(* IEC 61131-3 sources: Caravan/Archiv/12-04-19/Stations/Terminal/HMI/Network, 1 file *)

(* ---- ConfigObjects.st ---- *)
FUNCTION GLOBAL TAB TASK_CONF
_K_TASK, _K_REAL,
_K_END_VAR,

_K_TASK, _K_CYCLIC,
_K_END_VAR,

_K_TASK, _K_BACKGROUND,
_K_END_VAR,

_K_END_CONF
END_FUNCTION

FUNCTION GLOBAL TAB IPR_CONF
_K_IPR
	0$UINT,
_K_END_VAR,
_K_END_CONF
END_FUNCTION

FUNCTION GLOBAL TAB CONFIG_TABLES
00081$UINT,
0$UINT, 0, 10, "_ALARMDISPLAY",
0$UINT, 0, 11, "_ALARMX0PARA",
0$UINT, 0, 2, "_ALARMX1PARA",
0$UINT, 0, 19, "_ALARMXBUFFER",
0$UINT, 0, 1, "_BIT32",
0$UINT, 0, 1, "_BIT32RAM",
0$UINT, 0, 4, "_CAN",
0$UINT, 1, 3, "_CHECKONLINESTATUS",
0$UINT, 1, 0, "_CHECKSUM",
0$UINT, 1, 19, "_FILESYS",
0$UINT, 0, 14, "_GLOBAL",
0$UINT, 1, 2, "_GRAFIX",
0$UINT, 0, 1, "_HOTALARM",
0$UINT, 1, 8, "_IP",
0$UINT, 1, 1, "_IPCONFIGIF",
0$UINT, 1, 2, "_IPCONFIGMAIN",
0$UINT, 1, 2, "_IPCONFIGSTATION",
0$UINT, 0, 5, "_LANGUAGESELECTION",
0$UINT, 0, 1, "_LIMITMAX",
0$UINT, 0, 1, "_LIMITMIN",
0$UINT, 0, 114, "_LSE",
0$UINT, 1, 1, "_MULTITASK",
0$UINT, 0, 3, "_MYIO",
0$UINT, 0, 4, "_OSKERNEL",
0$UINT, 0, 6, "_OSZILSE",
0$UINT, 0, 0, "_OSZILSEBACKGROUND",
0$UINT, 0, 1, "_RADIO32",
0$UINT, 0, 1, "_RADIO32RAM",
0$UINT, 0, 3, "_SCREEN",
0$UINT, 0, 15, "_SCROLLAREA",
0$UINT, 0, 8, "_SCROLLAREA2",
0$UINT, 1, 0, "_SEARCHUSBFILETORESET",
0$UINT, 0, 0, "_STDLIB",
0$UINT, 2, 0, "_SYNCTIMEHMI",
0$UINT, 0, 7, "_SYSDATETIME",
0$UINT, 0, 0, "_SYSMSG",
0$UINT, 1, 1, "_TASKOBJECTCONTROL",
0$UINT, 1, 0, "_TOOLCAT",
0$UINT, 1, 1, "_WEATHERFORECAST",
0$UINT, 1, 0, "_WINDINDICATOR",
0$UINT, 0, 1, "_XACCESS",
0$UINT, 1, 4, "_XMLREADER",
0$UINT, 1, 2, "_XMLSTRUCTCREATOR",
0$UINT, 1, 7, "ALARMDISPLAYLIST",
0$UINT, 1, 1, "ALARMTITLELINE",
0$UINT, 1, 2, "CLIENT_SPLITTER_10",
0$UINT, 1, 1, "CLIENT_SPLITTER_BASE",
0$UINT, 0, 4, "CRITICALSECTION",
0$UINT, 1, 0, "DATAMANAGER",
0$UINT, 1, 0, "DATAMANAGERFIFO",
0$UINT, 1, 0, "DATAMANAGERPRIORITY",
0$UINT, 1, 37, "DISPLAYSETTINGS",
0$UINT, 0, 10, "GETBROADCASTDATA",
0$UINT, 0, 2, "GETTASKHANDLE",
0$UINT, 0, 1, "GRAPHIC",
0$UINT, 0, 0, "INPUTMYIO",
0$UINT, 2, 0, "KEYPADANUMSTDTEMPLATE",
0$UINT, 2, 0, "KEYPADIMAGESSTDTEMPLATE",
0$UINT, 1, 0, "KEYPADNUMSTDTEMPLATE",
0$UINT, 0, 0, "KOORDINATES_CLASS",
0$UINT, 1, 21, "MERKEREX",
0$UINT, 1, 31, "NETWORKCONFIG",
0$UINT, 1, 16, "PROJECTGLOBAL",
0$UINT, 1, 3, "RAM",
0$UINT, 1, 17, "RAMEX",
0$UINT, 1, 1, "RAMRINGBUFFER",
0$UINT, 1, 13, "SCREENSAVER",
0$UINT, 0, 23, "SIGCLIB",
0$UINT, 1, 10, "STRING",
0$UINT, 1, 82, "STRINGINTERNAL",
0$UINT, 1, 10, "STRINGRAM",
0$UINT, 0, 1, "SYSTEM",
0$UINT, 1, 5, "SYSTEMLOGGING",
0$UINT, 1, 14, "TCPCOMMUNICATION",
0$UINT, 1, 0, "TCPCOMMUNICATIONLOGFILTER",
0$UINT, 1, 4, "TCPCOMMUNICATIONLOGVIEWER",
0$UINT, 1, 3, "TITLELINE",
0$UINT, 1, 3, "TOUCHCALIB",
0$UINT, 1, 13, "USB_DATAEXCHANGE",
0$UINT, 1, 5, "USBDETECTION",
0$UINT, 1, 3, "VIRTUALBASEINIT",
ONE_CFG$UINT, 0, 0, "ONE_IPCONF_IPConfigHMI",
ONE_CFG$UINT, 0, 0, "ONE_Level_NET",
ONE_CFG$UINT, 0, 0, "ONE_LseRtkAlarm",
ONE_CFG$UINT, 0, 0, "ONE_LseRtkMain",
ONE_CFG$UINT, 1, 0, "ONE_NewAgeAlarmVis",
ONE_CFG$UINT, 1, 0, "ONE_NewAgeSettings",
ONE_CFG$UINT, 1, 0, "ONE_STDCommunicationToPLC",
ONE_CFG$UINT, 2, 0, "ONE_STDSettingsHMI",
ONE_CFG$UINT, 0, 0, "ONE_WEATHER_WeatherForecast",
TASK_CFG$UINT, 0, 0, "TASK_CONF",
IPR_CFG$UINT, 0, 0, "IPR_CONF",
PRJ_CFG$UINT, 0, 0, "HMI",
END_FUNCTION

#ifdef __LSLLDR_MULTIMASTER__
FUNCTION GLOBAL TAB CONFIG_MULTIMASTER
0000$UINT, 0001$UINT,
"MachineControl",
0005$UINT,
TO_UDINT(619908241), "SyncTimePLC.SyncDate", 0$USINT, 103$UINT, (0)$UDINT,
TO_UDINT(3791233966), "SyncTimePLC.SyncTime", 0$USINT, 103$UINT, (0)$UDINT,
TO_UDINT(4229011844), "Level_Class1.Level_Y_S", 0$USINT, 103$UINT, (0)$UDINT,
TO_UDINT(4258526131), "Level_Class1.Level_X_S", 0$USINT, 103$UINT, (0)$UDINT,
TO_UDINT(867522694), "_IPConfigIF1mc1.ClassSvr", 0$USINT, 103$UINT, (_MM_PROP_RO OR _MM_PROP_NEWINST)$UDINT,
END_FUNCTION
#endif

FUNCTION GLOBAL TAB CH_REDIRECT_EMB_TAB
0000$UINT,
00019$UINT,
"_WeatherForecast;Day1_DD_MM", "\Str_Day1_DD_MM.Data",
"_WeatherForecast;Day2_DD_MM", "\Str_Day2_DD_MM.Data",
"_WeatherForecast;Day3_DD_MM", "\Str_Day3_DD_MM.Data",
"_WeatherForecast;Day4_DD_MM", "\Str_Day4_DD_MM.Data",
"_WeatherForecast;Day5_DD_MM", "\Str_Day5_DD_MM.Data",
"_WeatherForecast;LastLocationName", "\Str_LastLocationName.Data",
"_WeatherForecast;ProxyAddress", "\Str_ProxyAddress.Data",
"_WeatherForecast;ProxyPassword", "\Str_ProxyPassword.Data",
"_WeatherForecast;ProxyPort", "\Str_ProxyPort.Data",
"_WeatherForecast;ProxyUser", "\Str_ProxyUser.Data",
"_WeatherForecast;WeatherLocCountry", "\Str_WeatherLocCountry.Data",
"_WeatherForecast;WeatherLocID", "\Str_WeatherLocID.Data",
"_WeatherForecast;WeatherLocName", "\Str_WeatherLocName.Data",
"_WeatherForecast;WeatherURL", "\Str_WeatherURL.Data",
"_WeatherForecast;WeatherUserID", "\Str_WeatherUserID.Data",
"AlarmDisplayList;AlaTxtLong", "\AlarmTxtLong.Data",
"AlarmDisplayList;AlaTxtShort", "\AlarmTxtShort.Data",
"TCPCommunication;TaskName", "\ThreadName.Data",
"USBDetection;DriveLetter", "\USBDriveLetter.Data",
END_FUNCTION
